FUNCTION_BLOCK FB_RelayMonostable IMPLEMENTS I_Relay
VAR_INPUT
    stDeviceId : ST_DeviceId;
END_VAR
VAR_OUTPUT
    bOutput : BOOL;
END_VAR
VAR
    bRequestedState : BOOL;
END_VAR

bOutput := bRequestedState;

PROPERTY DeviceId : ST_DeviceId
GET
DeviceId := stDeviceId;
END_GET
END_PROPERTY

PROPERTY IsOn : BOOL
GET
IsOn := bOutput;
END_GET
END_PROPERTY

METHOD PUBLIC TurnOn
bRequestedState := TRUE;
END_METHOD

METHOD PUBLIC TurnOff
bRequestedState := FALSE;
END_METHOD

METHOD PUBLIC Toggle
bRequestedState := NOT bRequestedState;
END_METHOD

END_FUNCTION_BLOCK

(* stored: Version 1.1.0.1, ProductVersion 3.1.4026.20
   POU FB_RelayMonostable: Id {66666666-6666-4666-8666-666666666660}
   Property DeviceId: Id {66666666-6666-4666-8666-666666666661}
   Get Get: Id {66666666-6666-4666-8666-666666666671}
   Property IsOn: Id {66666666-6666-4666-8666-666666666662}
   Get Get: Id {66666666-6666-4666-8666-666666666672}
   Method TurnOn: Id {66666666-6666-4666-8666-666666666663}
   Method TurnOff: Id {66666666-6666-4666-8666-666666666664}
   Method Toggle: Id {66666666-6666-4666-8666-666666666665} *)
